(*
SPDX-FileCopyrightText: © 2026 Oleksandr Tiutyk <trofimich@gmail.com>
SPDX-License-Identifier: MIT
License: https://opensource.org/license/mit
*)

(*!
<summary>
Beckhoff bidirectional strain gauge / resistor bridge channel process image.
</summary>
<description>
Aggregates input status/value (STRAIN_GAUGE_INPUT_CHANNEL) and output control (STRAIN_GAUGE_OUTPUT_CHANNEL)
for one measuring bridge channel.
When used for I/O, link located fields or their containing buffers to the matching selected PDOs.
The record is not a packed wire buffer; compiler padding is not part of the device specification.
Unlinked/default values do not prove valid I/O. The caller evaluates bus/channel validity before use.
Use one owner task per instance and externally synchronize other access; multi-field snapshots are not atomic.
Copies store data without creating hardware links. Keep borrowed field references valid while consumers are bound.
This passive record performs no validation, synchronization, configuration or protocol advancement.
</description>
*)
TYPE STRAIN_GAUGE_CHANNEL :
STRUCT
	In : STRAIN_GAUGE_INPUT_CHANNEL;
	Out : STRAIN_GAUGE_OUTPUT_CHANNEL;
END_STRUCT
END_TYPE

(* stored: Version 1.1.0.1, ProductVersion 3.1.4026.20
   DUT STRAIN_GAUGE_CHANNEL: Id {5dac29e2-5891-4a4d-aa11-27f72e8de5ae} *)
